// Raw analog value to engineering units
FUNCTION F_Old : REAL
VAR_INPUT
	nRaw : INT;
	fMax : REAL;
END_VAR
VAR
	fTmp : REAL;
END_VAR

fTmp := INT_TO_REAL(nRaw) / 32767.0;
F_Old := fTmp * fMax;

END_FUNCTION

(* stored: Version 1.1.0.1, ProductVersion 3.1.4026.12
   POU F_Old: Id {3a2b3c4d-0000-4000-8000-000000000003}, SpecialFunc None *)
